(* IEC 61131-3 sources: PLC_Gen_Frame/Agents4PLC_release/results/task_1778477714, 1 file *)

(* ---- output.ST ---- *)
FUNCTION_BLOCK AGVControlSystem
VAR_INPUT
    MaterialRequest : INT;
END_VAR
VAR_OUTPUT
    AGV1_Ready : BOOL;
    AGV2_Ready : BOOL;
    AGV3_Ready : BOOL;
END_VAR

// Generated by DummyPLCGenerator

END_FUNCTION_BLOCK
